(*
SPDX-FileCopyrightText: c 2026 Oleksandr Tiutyk <trofimich@gmail.com>
SPDX-License-Identifier: MIT
License: https://opensource.org/license/mit
*)

(*!
<summary>Checks direct analog output processing for a bound INT16 value.</summary>
<description>
Uses a live case-owned automation parent and fresh local device fixtures on every run.
The scenario reads and writes ordinary simulated storage within one task cycle.
</description>
*)

{attribute 'no_assign'}
{attribute 'no_explicit_call' := 'do not call this function block directly'}
FUNCTION_BLOCK AnalogOutputScalingTest EXTENDS TOF_Testing.SingleCycleTest
VAR_STAT
	{attribute 'hide'}
	_ClassName : STRING := __POUNAME();
END_VAR
VAR
	//! <summary>Live parent borrowed by the method-local simulated device.</summary>
	_AutomationRoot : MockAutomationController(name := "DevicesIORoot");
END_VAR

(*!
<summary>Checks direct analog output processing for a bound INT16 value.</summary>
*)
METHOD PROTECTED ExecuteTest
VAR
	converter : TOF_Devices_IO.DirectAnalogValueConverter;
	analogOutput : TOF_Devices_IO.AnalogOutput(name := "AO_Test", parent := _AutomationRoot, converter := converter);
	rawOutput : INT;
END_VAR
analogOutput.Initialize();
analogOutput.BindToInt16IO(rawVariable := rawOutput);

analogOutput.Value := 750.0;
analogOutput.ProcessOutput();

Assert.ThatInt(
	actual := rawOutput,
	message := "Raw INT output should match 750"
).ToBe(expected := 750);
END_METHOD

//! <summary>Borrows the concrete class name. Callers must not modify it.</summary>
{attribute 'monitoring' := 'call'}
PROPERTY ClassName : REFERENCE TO STRING
GET
ClassName REF= _ClassName;
END_GET
END_PROPERTY

//! <summary>Borrows the compiler-initialized namespace name. Callers must not modify it.</summary>
{attribute 'monitoring' := 'call'}
PROPERTY NamespaceName : REFERENCE TO STRING
GET
NamespaceName REF= CurrentNamespace.Name;
END_GET
END_PROPERTY

//! <summary>Reports the concrete instance size in bytes.</summary>
{attribute 'monitoring' := 'call'}
PROPERTY SelfSize : ULINT
GET
SelfSize := XSIZEOF(THIS^);
END_GET
END_PROPERTY

END_FUNCTION_BLOCK

(* stored: Version 1.1.0.1
   POU AnalogOutputScalingTest: Id {4ace37ab-816c-4339-abb9-aa1d155852c4}, SpecialFunc None
   Method ExecuteTest: Id {16723a4b-4261-459b-8403-90317d1668ed}
   Property ClassName: Id {21c8e7e4-fd39-4de5-95c7-b70de6980f16}
   Get Get: Id {3ba647c5-acbc-4cd4-895e-075b0c88aed0}
   Property NamespaceName: Id {313841be-7ada-49d8-9970-db5914e2cfbc}
   Get Get: Id {783907fd-dad6-4a52-a118-a1ca46950546}
   Property SelfSize: Id {5221818f-89ef-45a6-8d39-a163041dde48}
   Get Get: Id {d9785026-c99e-4167-9cb5-61052fbf0334} *)
